(* IEC 61131-3 sources: Test-Git_ESME26/TestProgettoESME_26.fbsproj/AxisModule_Migration_Example.device.xml.v3^/Plc Logic.plclogic.xml.v3^/Application.application.xml.v3^/Sercos_AxisModule, 2 files *)

(* ---- FB_Set230VModeAsync.fb.st ---- *)
FUNCTION_BLOCK FB_Set230VModeAsync IMPLEMENTS SE_Async.IF_Async
VAR_INPUT
	i_ifSercosIdentificationAccess : SDI.IF_SercosIdentificationAccess;
END_VAR
VAR_OUTPUT
	q_diResult : DINT;
	q_sDiagMsg : STRING[255];
END_VAR
VAR
	xDone_loc : Bool;
END_VAR

(* ---- SR_Sercos.prg.st ---- *)
PROGRAM SR_Sercos

VAR_OUTPUT
	q_xSercosRun: BOOL;
END_VAR
// configuration
VAR
	fbSet230VModeAsync	: FB_Set230VModeAsync;
 	etMainsVoltageMode : ET_MainsVoltageMode := ET_MainsVoltageMode._230V;
END_VAR

VAR
	xInit : BOOL := TRUE;
	xResetSercos: BOOL;
	bDiagQuit :BOOL := FALSE;
    diState :DINT:=0;
	xError: BOOL;
	etResult: MOIN.ET_Result;
	xError2: BOOL;
	etResult2: MOIN.ET_Result;

	diResult : DINT;
	sDiagMsg : STRING[255];

END_VAR

CASE diState OF
	0:
		IF xInit THEN
			IF PSM_Lexium62.WorkingMode.DesiredMode = CFDI.ET_WorkingMode.Virtual THEN
				diState := 70;
			ELSE
				diState := 20;
			END_IF
		END_IF
	20:
		SE_Async.G_ifAsyncMgr.Init();
		IF SE_Async.G_ifAsyncMgr.xInitDone THEN
			// go to CP2
			SercosMaster.SercosPhaseChanger.DesiredPhase := SMI.ET_SercosPhase.Phase2;
			diState                                      := diState + 10;
		END_IF

	30:
		// wait for CP2
		IF SercosMaster.SercosPhaseChanger.ActualState = SMI.ET_SercosState.Phase2 THEN
			diState := diState + 10;
		END_IF

	40:
		// configure 230V mode on PowerSupply
		IF etMainsVoltageMode = ET_MainsVoltageMode._230V THEN
			fbSet230VModeAsync(i_ifSercosIdentificationAccess := PSM_Lexium62);
			fbSet230VModeAsync.xDone := FALSE;
			SE_Async.G_ifAsyncMgr.Start(fbSet230VModeAsync);
			diState := diState + 10;
		ELSE
			diState := 70;
		END_IF

	50:
		// configure 230V mode on DRV_Slave1
		IF fbSet230VModeAsync.xDone THEN
			fbSet230VModeAsync(i_ifSercosIdentificationAccess := DRV_Slave1);
			fbSet230VModeAsync.xDone := FALSE;
			SE_Async.G_ifAsyncMgr.Start(fbSet230VModeAsync);
			diState := diState + 10;
		ELSIF fbSet230VModeAsync.q_diResult <> 0 THEN
			sDiagMsg := fbSet230VModeAsync.q_sDiagMsg;
			diState  := 500;
			RETURN;
		END_IF

	60:
		// configure 230V mode on DRV_Slave2
		IF fbSet230VModeAsync.xDone THEN
			fbSet230VModeAsync(i_ifSercosIdentificationAccess := DRV_Slave2);
			fbSet230VModeAsync.xDone := FALSE;
			SE_Async.G_ifAsyncMgr.Start(fbSet230VModeAsync);
			diState := diState + 10;
		ELSIF fbSet230VModeAsync.q_diResult <> 0 THEN
			sDiagMsg := fbSet230VModeAsync.q_sDiagMsg;
			diState  := 500;
			RETURN;
		END_IF

	70:
		// go to CP4
		SercosMaster.SercosPhaseChanger.DesiredPhase := SMI.ET_SercosPhase.Phase4;
		diState                                      := diState + 10;
	80:
		// wait for CP4
		IF SercosMaster.SercosPhaseChanger.ActualState = SMI.ET_SercosState.Phase4 THEN
			diState      := diState + 10;
			q_xSercosRun := TRUE;
		END_IF
	90:
		IF xResetSercos THEN
			xResetSercos 								 := FALSE;
			q_xSercosRun                                 := FALSE;
			SercosMaster.SercosPhaseChanger.DesiredPhase := SMI.ET_SercosPhase.NRT;
			diState                                      := 0;
		END_IF
END_CASE

IF bDiagQuit THEN
	bDiagQuit := FALSE;
	SEC.FC_DiagAcknowledge();
END_IF
